// TIA Portal V20 export
Screen "Valve8Pos"  1276x673
  ScreenItem "OBJECT_37" at 2,226 size 635x25  Type=HmiTextBox
  ScreenItem "OBJECT_40" at 642,96 size 635x25  Type=HmiTextBox
  ScreenItem "OBJECT_42" at 642,70 size 635x25  Type=HmiTextBox
  ScreenItem "OBJECT_47" at 642,174 size 635x25  Type=HmiTextBox
  ScreenItem "OBJECT_48" at 642,226 size 635x25  Type=HmiTextBox
  ScreenItem "OBJECT_51" at 642,252 size 635x25  Type=HmiTextBox
  ScreenItem "OBJECT_15" at 2,252 size 635x25  Type=HmiTextBox
  ScreenItem "OBJECT_24" at 2,278 size 635x25  Type=HmiTextBox
  ScreenItem "OBJECT_27" at 2,356 size 635x25  Type=HmiTextBox
  ScreenItem "OBJECT_28" at 2,382 size 635x25  Type=HmiTextBox
  ScreenItem "OBJECT_30" at 2,122 size 635x25  Type=HmiTextBox
  ScreenItem "OBJECT_31" at 2,96 size 635x25  Type=HmiTextBox
  ScreenItem "OBJECT_33" at 2,174 size 635x25  Type=HmiTextBox
  ScreenItem "OBJECT_34" at 2,148 size 635x25  Type=HmiTextBox
  ScreenItem "OBJECT_35" at 2,200 size 635x25  Type=HmiTextBox
  ScreenItem "OBJ1" at 642,122 size 635x25  Type=HmiTextBox
  ScreenItem "OBJECT_2" at 642,148 size 635x25  Type=HmiTextBox
  ScreenItem "OBJECT_3" at 642,200 size 635x25  Type=HmiTextBox
  ScreenItem "OBJECT_4" at 642,278 size 635x25  Type=HmiTextBox
  ScreenItem "OBJECT_5" at 642,304 size 635x25  Type=HmiTextBox
  ScreenItem "Title_ScreenOverview_X390_Y2" at 687,5 size 144x30  Type=HmiSymbolicIOField
  ScreenItem "OBJECT_1" at 2,330 size 635x25  Type=HmiTextBox
  ScreenItem "OBJECT_6" at 2,304 size 635x25  Type=HmiTextBox
  ScreenItem "TecUnit_Type" at 571,35 size 200x22  Type=HmiTextBox
  ScreenItem "Line_Header_X0_Y64" at 0,64 size 1276x0  Type=HmiLine
  ScreenItem "Reserved_2" at 642,330 size 635x25  Type=HmiTextBox
  ScreenItem "Textfield_Overview_Alarms" at 910,32 size 100x25  Type=HmiTextBox
  ScreenItem "Tec-Unit-Diag_Legend" at 1184,2 size 90x60  Type=HmiButton
  ScreenItem "OBJECT_7" at 2,70 size 635x25  Type=HmiTextBox
  ScreenItem "Position_Left_9" at 10,542 size 45x20  Type=HmiTextBox
  ScreenItem "Position_Left_10" at 10,498 size 45x20  Type=HmiTextBox
  ScreenItem "Screen_Back_X0-Y65-W1280-H585" at 0,69 size 1280x581  Type=HmiButton
  ScreenItem "Position_Left_11" at 10,520 size 45x20  Type=HmiTextBox
  ScreenItem "Grafik_Cylinder_23" at 1150,470 size 60x112  Type=HmiGraphicView
  ScreenItem "Position_Left_8" at 1164,542 size 30x20  Type=HmiTextBox
  ScreenItem "Position_Right_8" at 1164,498 size 30x20  Type=HmiTextBox
  ScreenItem "Position_Y8" at 1164,520 size 30x20  Type=HmiTextBox
  ScreenItem "Text_Cylinder_23" at 1156,474 size 50x21  Type=HmiTextBox
  ScreenItem "Grafik_Cylinder_22" at 995,470 size 60x112  Type=HmiGraphicView
  ScreenItem "Position_Left_7" at 1009,542 size 30x20  Type=HmiTextBox
  ScreenItem "Position_Right_7" at 1009,498 size 30x20  Type=HmiTextBox
  ScreenItem "Position_Y7" at 1009,520 size 30x20  Type=HmiTextBox
  ScreenItem "Text_Cylinder_22" at 1001,474 size 50x21  Type=HmiTextBox
  ScreenItem "Grafik_Cylinder_21" at 841,471 size 60x112  Type=HmiGraphicView
  ScreenItem "Position_Left_6" at 855,542 size 30x20  Type=HmiTextBox
  ScreenItem "Position_Right_6" at 855,498 size 30x20  Type=HmiTextBox
  ScreenItem "Position_Y6" at 855,520 size 30x20  Type=HmiTextBox
  ScreenItem "Text_Cylinder_21" at 847,475 size 50x21  Type=HmiTextBox
  ScreenItem "Grafik_Cylinder_20" at 687,470 size 60x112  Type=HmiGraphicView
  ScreenItem "Position_Left_5" at 701,542 size 30x20  Type=HmiTextBox
  ScreenItem "Position_Right_5" at 701,498 size 30x20  Type=HmiTextBox
  ScreenItem "Position_Y5" at 701,520 size 30x20  Type=HmiTextBox
  ScreenItem "Text_Cylinder_20" at 693,474 size 50x21  Type=HmiTextBox
  ScreenItem "Grafik_Cylinder_19" at 532,470 size 60x112  Type=HmiGraphicView
  ScreenItem "Position_Left_4" at 546,542 size 30x20  Type=HmiTextBox
  ScreenItem "Position_Right_4" at 546,498 size 30x20  Type=HmiTextBox
  ScreenItem "Position_Y4" at 546,520 size 30x20  Type=HmiTextBox
  ScreenItem "Text_Cylinder_19" at 538,474 size 50x21  Type=HmiTextBox
  ScreenItem "Grafik_Cylinder_18" at 378,470 size 60x112  Type=HmiGraphicView
  ScreenItem "Position_Left_3" at 392,542 size 30x20  Type=HmiTextBox
  ScreenItem "Position_Right_3" at 392,498 size 30x20  Type=HmiTextBox
  ScreenItem "Position_Y3" at 392,520 size 30x20  Type=HmiTextBox
  ScreenItem "Text_Cylinder_18" at 384,474 size 50x21  Type=HmiTextBox
  ScreenItem "Grafik_Cylinder_17" at 224,470 size 60x112  Type=HmiGraphicView
  ScreenItem "Position_Left_2" at 238,542 size 30x20  Type=HmiTextBox
  ScreenItem "Position_Right_2" at 238,498 size 30x20  Type=HmiTextBox
  ScreenItem "Position_Y2" at 238,520 size 30x20  Type=HmiTextBox
  ScreenItem "Text_Cylinder_17" at 230,474 size 50x21  Type=HmiTextBox
  ScreenItem "Grafik_Cylinder_16" at 101,467 size 60x112  Type=HmiGraphicView
  ScreenItem "Position_Right_1" at 115,495 size 30x20  Type=HmiTextBox
  ScreenItem "Position_Left_1" at 115,539 size 30x20  Type=HmiTextBox
  ScreenItem "Position_Y1" at 115,517 size 30x20  Type=HmiTextBox
  ScreenItem "Text_Cylinder_16" at 107,471 size 50x21  Type=HmiTextBox
  ScreenItem "Title_ScreenOverview_X390_Y2_1" at 511,5 size 162x30  Type=HmiSymbolicIOField
  ScreenItem "permanentareaborderrectangle" at 0,0 size 0x0  Type=HmiRectangle
  ScreenItem "Button_Back" at 2,2 size 90x60  Type=HmiButton
  ScreenItem "Textfield_Overview_State_1" at 284,32 size 100x25  Type=HmiTextBox
